Fanuc KAREL source: KT00782.KL

PROGRAM KT00782
%NOLOCKGROUP
VAR
  S1: STRING[80]
  S2: STRING[80]
  OUT: INTEGER
BEGIN
  S1 = 'A'
  S2 = 'B'
  S1 = 'A'
  S2 = 'B'
  OUT = ASIN(S1)
END KT00782
